TYPE Shuttle_Position_UDT :
STRUCT
	x: DINT;
	y: DINT;
	Charging: BOOL;
END_STRUCT
END_TYPE

(* stored: Version 1.1.0.1
   DUT Shuttle_Position_UDT: Id {31406683-9a9e-47a2-ad9e-671dbded8aac} *)
